// Generic 1 kHz motion-profile generator for the V3.2 motor. Evaluates the
// selected shape as value(t) online (no precomputed array) and streams it to
// the field PRG_Motion routes by nField. Shapes ported from the Cheetah
// ProfileGenerator: Sinusoidal / Trapezoidal / Step / S-Curve / Ramp, plus
// two point-to-point shapes (velocity-trapezoid displacement, planned by the
// app from v_max/a_max): P2P moves one leg and holds at the end; P2P_RT goes
// out and back (v = 0 at the turnaround), so repetitive reps chain without a
// jump. For both, fPeakValue is the SIGNED cruise velocity, fAccelTime/
// fSteadyTime/fDecelTime are the leg's segment times, and fStartValue is the
// ABSOLUTE anchor position the app planned from (exact landing on target).
//
// On Start the command is LATCHED into 'cfg' (a local copy of stTraj). The
// generator + the valueAt method read 'cfg' only -- so mid-run parameter
// changes are ignored, and the method never touches the VAR_IN_OUT (no C0371).
//
// Anchoring: for position-target fields (nField 0/1) the profile rides on the
// rotor's position captured at Start -> out = startPos + (value(t) - value(0)),
// so it begins exactly where the motor is (no jump). Velocity/current (2/3) use
// the value directly. Repetitive loops the whole profile (nReps; 0 = infinite),
// resting fRestS between reps.
FUNCTION_BLOCK FB_TrajectoryGen
VAR_IN_OUT
    stTraj          : ST_MenteeTrajCmd;
END_VAR
VAR_INPUT
    fMeasuredPos    : REAL;     // current measured output position [rad]
    fDt             : REAL;     // task cycle time [s]
    bStartSync      : BOOL;     // shared synchronized start (PRG_Motion gates with the Mentee enable)
    bStopSync       : BOOL;     // shared synchronized stop
END_VAR
VAR_OUTPUT
    bRunning        : BOOL;
    fSetpoint       : REAL;
    nFieldOut       : BYTE;     // LATCHED field of the running profile — route by
                                // this, not the live stTraj.nField, so an ADS
                                // reconfig mid-run can't misroute the output
END_VAR
VAR
    cfg             : ST_MenteeTrajCmd;   // latched command (read by body + valueAt)
    rStart          : R_TRIG;
    rStop           : R_TRIG;
    eState          : INT;      // see ST_* constants
    fElapsed        : REAL;     // time into the current run [s]
    fTotalDur       : REAL;     // total duration of one run [s]
    fStartPos       : REAL;     // anchor position (captured at Start)
    fValue0         : REAL;     // value(0) for anchoring
    bAnchor         : BOOL;     // position-target field -> anchor at current pos
    nRepDone        : UDINT;
    fRest           : REAL;     // rest countdown [s]
    fRaw            : REAL;
    bWasActive      : BOOL;
END_VAR
VAR CONSTANT
    ST_IDLE         : INT := 0;
    ST_RUN          : INT := 1;
    ST_REST         : INT := 2;
    ST_DONE         : INT := 3;
    SH_SINE         : BYTE := 0;
    SH_TRAP         : BYTE := 1;
    SH_STEP         : BYTE := 2;
    SH_SCURVE       : BYTE := 3;
    SH_RAMP         : BYTE := 4;
    SH_P2P          : BYTE := 5;
    SH_P2P_RT       : BYTE := 6;
END_VAR

rStart(CLK := stTraj.bStart OR bStartSync);
rStop(CLK := stTraj.bStop OR bStopSync);

// Stop -> hold current position (idle; PRG_Motion stops overriding the field).
IF rStop.Q THEN
    eState := ST_IDLE;
END_IF

// Start a new run -> latch the command into cfg; everything below reads cfg.
IF rStart.Q AND (stTraj.nShape <= SH_P2P_RT) AND (stTraj.nField <= 3) THEN
    cfg      := stTraj;
    nFieldOut := cfg.nField;
    fElapsed := 0.0;
    nRepDone := 0;
    // P2P ends AWAY from its start, so replaying it would jump the setpoint
    // back -> one-way moves are never repetitive (oscillation uses SH_P2P_RT).
    IF cfg.nShape = SH_P2P THEN
        cfg.bRepetitive := FALSE;
    END_IF
    // total duration of one run, per shape
    IF (cfg.nShape = SH_TRAP) OR (cfg.nShape = SH_SCURVE) OR (cfg.nShape = SH_P2P) THEN
        fTotalDur := cfg.fAccelTime + cfg.fSteadyTime + cfg.fDecelTime;
    ELSIF cfg.nShape = SH_P2P_RT THEN
        fTotalDur := 2.0 * (cfg.fAccelTime + cfg.fSteadyTime + cfg.fDecelTime);
    ELSE
        fTotalDur := cfg.fDuration;
    END_IF
    // position-target fields ride on the current position (no jump). The P2P
    // shapes anchor on the app's PLANNED start (fStartValue) instead, so the
    // move lands EXACTLY on the planned target; any drift accrued since
    // planning shows as a small initial step the servo absorbs (identical to
    // the app-side streamer these shapes replace).
    bAnchor := (cfg.nField = 0) OR (cfg.nField = 1);
    IF bAnchor THEN
        IF (cfg.nShape = SH_P2P) OR (cfg.nShape = SH_P2P_RT) THEN
            fStartPos := cfg.fStartValue;
        ELSE
            fStartPos := fMeasuredPos;
        END_IF
        fValue0   := valueAt(0.0);
    ELSE
        fStartPos := 0.0;
        fValue0   := 0.0;
    END_IF
    eState := ST_RUN;
END_IF

// "Active this cycle" is latched BEFORE transitions so the cycle that ends the
// run still writes the final value.
bWasActive := (eState = ST_RUN) OR (eState = ST_REST);

CASE eState OF

ST_RUN:
    fRaw := valueAt(fElapsed);
    IF bAnchor THEN
        stTraj.fSetpoint := fStartPos + (fRaw - fValue0);
    ELSE
        stTraj.fSetpoint := fRaw;
    END_IF
    fElapsed := fElapsed + fDt;
    IF fElapsed >= fTotalDur THEN
        // land on the exact end value
        fRaw := valueAt(fTotalDur);
        IF bAnchor THEN
            stTraj.fSetpoint := fStartPos + (fRaw - fValue0);
        ELSE
            stTraj.fSetpoint := fRaw;
        END_IF
        IF NOT cfg.bRepetitive THEN
            eState := ST_DONE;
        ELSE
            nRepDone := nRepDone + 1;
            IF (cfg.nReps > 0) AND (nRepDone >= cfg.nReps) THEN
                eState := ST_DONE;
            ELSE
                fRest  := cfg.fRestS;
                eState := ST_REST;
            END_IF
        END_IF
    END_IF

ST_REST:
    fRest := fRest - fDt;                   // hold last setpoint during the rest
    IF fRest <= 0.0 THEN
        fElapsed := 0.0;
        eState   := ST_RUN;
    END_IF

ST_DONE:
    ;                                       // hold fSetpoint

ST_IDLE:
    ;                                       // not running

END_CASE

stTraj.fElapsed := fElapsed;
bRunning        := bWasActive;
fSetpoint       := stTraj.fSetpoint;
stTraj.bRunning := bRunning;

// Signed displacement along one point-to-point velocity-trapezoid leg at
// time fT [s]: accelerate 0 -> fPeakValue over fAccelTime, cruise for
// fSteadyTime, decelerate back to 0 over fDecelTime. Clamps past the end, so
// leg(end) = fPeakValue * (fAccelTime/2 + fSteadyTime + fDecelTime/2) = the
// leg distance. Mirrors the app's TrapezoidProfile (trajectory.py) exactly.
METHOD p2pLeg : REAL
VAR_INPUT
    fT  : REAL;
END_VAR
VAR
    fTa : REAL;     // accel time [s]
    fTc : REAL;     // cruise time [s]
    fTd : REAL;     // decel time [s]
    fV  : REAL;     // signed cruise velocity
    fU  : REAL;
END_VAR
fTa := MAX(cfg.fAccelTime, 1E-6);
fTc := cfg.fSteadyTime;
fTd := MAX(cfg.fDecelTime, 1E-6);
fV  := cfg.fPeakValue;

IF fT <= 0.0 THEN
    p2pLeg := 0.0;
ELSIF fT < fTa THEN
    // accelerating: 1/2 * a * t^2 with a = fV / fTa
    p2pLeg := 0.5 * fV * fT * fT / fTa;
ELSIF fT < (fTa + fTc) THEN
    // cruising
    p2pLeg := fV * (0.5 * fTa + (fT - fTa));
ELSE
    // decelerating (clamped at the leg end)
    fU := fT - fTa - fTc;
    IF fU > fTd THEN fU := fTd; END_IF
    p2pLeg := fV * (0.5 * fTa + fTc + fU - 0.5 * fU * fU / fTd);
END_IF
END_METHOD

// Shape value at time fT [s] — closed-form, mirrors the Cheetah ProfileGenerator.
// Reads the latched 'cfg' (FB-local), never the VAR_IN_OUT.
METHOD valueAt : REAL
VAR_INPUT
    fT  : REAL;
END_VAR
VAR
    fU  : REAL;
END_VAR
VAR CONSTANT
    TWO_PI : REAL := 6.2831853;
END_VAR
CASE cfg.nShape OF

0:  // Sinusoidal: offset + A * sin(2*pi*f*t)
    valueAt := cfg.fOffset + cfg.fAmplitude * SIN(TWO_PI * cfg.fFrequency * fT);

1:  // Trapezoidal: ramp start->peak / hold / ramp peak->start
    IF fT < cfg.fAccelTime THEN
        valueAt := cfg.fStartValue
                 + (cfg.fPeakValue - cfg.fStartValue) * (fT / MAX(cfg.fAccelTime, 1E-6));
    ELSIF fT < (cfg.fAccelTime + cfg.fSteadyTime) THEN
        valueAt := cfg.fPeakValue;
    ELSE
        fU := (fT - cfg.fAccelTime - cfg.fSteadyTime) / MAX(cfg.fDecelTime, 1E-6);
        IF fU > 1.0 THEN fU := 1.0; END_IF
        valueAt := cfg.fPeakValue - (cfg.fPeakValue - cfg.fStartValue) * fU;
    END_IF

2:  // Step: start until step time, then end
    IF fT < cfg.fStepTime THEN
        valueAt := cfg.fStartValue;
    ELSE
        valueAt := cfg.fEndValue;
    END_IF

3:  // S-Curve: quintic smoothstep start->peak / hold / peak->start
    IF fT < cfg.fAccelTime THEN
        fU := fT / MAX(cfg.fAccelTime, 1E-6);
        valueAt := cfg.fStartValue
                 + (cfg.fPeakValue - cfg.fStartValue) * (fU*fU*fU*(10.0 + fU*(-15.0 + fU*6.0)));
    ELSIF fT < (cfg.fAccelTime + cfg.fSteadyTime) THEN
        valueAt := cfg.fPeakValue;
    ELSE
        fU := (fT - cfg.fAccelTime - cfg.fSteadyTime) / MAX(cfg.fDecelTime, 1E-6);
        IF fU > 1.0 THEN fU := 1.0; END_IF
        valueAt := cfg.fPeakValue
                 - (cfg.fPeakValue - cfg.fStartValue) * (fU*fU*fU*(10.0 + fU*(-15.0 + fU*6.0)));
    END_IF

4:  // Ramp: linear start->end over duration
    fU := fT / MAX(cfg.fDuration, 1E-6);
    IF fU > 1.0 THEN fU := 1.0; END_IF
    valueAt := cfg.fStartValue + (cfg.fEndValue - cfg.fStartValue) * fU;

5:  // P2P: one-way velocity-trapezoid displacement; ends at the leg distance
    valueAt := p2pLeg(fT);

6:  // P2P round trip: leg out, then the same leg mirrored back to the start
    fU := cfg.fAccelTime + cfg.fSteadyTime + cfg.fDecelTime;   // one leg [s]
    IF fT < fU THEN
        valueAt := p2pLeg(fT);
    ELSE
        valueAt := p2pLeg(fU) - p2pLeg(fT - fU);
    END_IF

ELSE
    valueAt := 0.0;
END_CASE
END_METHOD

END_FUNCTION_BLOCK

(* stored: Version 1.1.0.1, ProductVersion 3.1.4026.18
   POU FB_TrajectoryGen: Id {c2f8d1b3-5e42-4a7b-8d3f-6b1c2e3a4d50}, SpecialFunc None
   Method p2pLeg: Id {a7c4e5f6-2b83-4d1a-9c5e-8f3a4b6d7e92}
   Method valueAt: Id {d3a9e2c4-6f53-4b8c-9e4a-7c2d3f4b5e61} *)
